{attribute 'qualified_only'}
{attribute 'strict'}
TYPE E_Filling_State :
(
	eNot_Ready := 0,
	eReady_ToFill,
	eFilling_InProcess
);
END_TYPE

(* stored: Version 1.1.0.1, ProductVersion 3.1.4024.15
   DUT E_Filling_State: Id {219e501c-0109-47a4-973b-411e6e86c6c0} *)
